// État d'une alarme active (docs/14 § 5)
{attribute 'qualified_only'}
{attribute 'strict'}
TYPE E_AlarmState :
(
    ActiveUnacked := 0,
    ActiveAcked := 1,
    ClearedUnacked := 2
) USINT;
END_TYPE

(* stored: Version 1.1.0.1, ProductVersion 3.1.4024.12
   DUT E_AlarmState: Id {ec99e4ab-e67e-5945-8e15-4bc5055c19a1} *)
